(* IEC 61131-3 sources: Caravan/Archiv/12-04-19/Stations/Terminal/HMI/Class/_WeatherForecast (part 2) *)

  for i:=0 to (StrLength - 1) do
    if ((myBuffer[BufferPos - i] >= '0') & (myBuffer[BufferPos - i] <= '9')) then
      case i of
        0: RetValue += TO_DINT((myBuffer[BufferPos - i] - '0') * 1);
        1: RetValue += TO_DINT((myBuffer[BufferPos - i] - '0') * 10);
        2: RetValue += TO_DINT((myBuffer[BufferPos - i] - '0') * 100);
        3: RetValue += TO_DINT((myBuffer[BufferPos - i] - '0') * 1000);
        4: RetValue += TO_DINT((myBuffer[BufferPos - i] - '0') * 10000);
        5: RetValue += TO_DINT((myBuffer[BufferPos - i] - '0') * 100000);
        6: RetValue += TO_DINT((myBuffer[BufferPos - i] - '0') * 1000000);
        7: RetValue += TO_DINT((myBuffer[BufferPos - i] - '0') * 10000000);
        8: RetValue += TO_DINT((myBuffer[BufferPos - i] - '0') * 100000000);
        9: RetValue += TO_DINT((myBuffer[BufferPos - i] - '0') * 1000000000);
      end_case;

    elsif (myBuffer[BufferPos - i] = '-') then    // negate
      RetValue := RetValue * -1;
    elsif ((myBuffer[BufferPos - i] = '.') | (myBuffer[BufferPos - i] = ',')) then    // start again in case of comma
      if ((myBuffer[BufferPos - i+1] - '0') >= 5) then
        RetValue := 1;
      else
        RetValue := 0;
      end_if;
      StrLength -= (i+1);
      i := -1;
      BufferPos := StrLength - 1;
    end_if;

  end_for;

END_FUNCTION

FUNCTION _WeatherForecast::MakeLocalTime
	VAR_INPUT
		pInTime 	: ^CHAR;
		UTC_Offset 	: DINT;
		pRetTime 	: ^CHAR;
	END_VAR

  VAR
  	myTime    : SYSTIME;
  	myDate    : SYSDATE;
    unixtime    : UDINT;
    myTxt : ARRAY [0..20] OF USINT;
  END_VAR

  if ((pInTime <> NIL) & (pRetTime <> NIL)) then

    myTime.wHour   := TO_UINT(CharToDint(pInTime +11, DataLen:=2));
    myTime.wMinute := TO_UINT(CharToDint(pInTime +14, DataLen:=2));
    myTime.wSecond := TO_UINT(CharToDint(pInTime +17, DataLen:=2));
    myTime.wSecond += 1;  // KaiAnd: workaround against UnixTimeStampConvert() bug (2017-10-01 00:00:00 -> 2017-09-31 00:00:00)

    myDate.wYear  := TO_UINT(CharToDint(pInTime +0, DataLen:=4));
    myDate.wMonth := TO_UINT(CharToDint(pInTime +5, DataLen:=2));
    myDate.wDay   := TO_UINT(CharToDint(pInTime +8, DataLen:=2));

    unixtime := SigCLib.UnixTimeStampReconvert(#myDate, #myTime);

    if (UTC_Offset > 0) then
      unixtime += TO_UDINT(UTC_Offset*3600);
    else
      unixtime -= TO_UDINT(UTC_Offset*-1 *3600);
    end_if;

    SigCLib.UnixTimeStampConvert(#myDate, #myTime, unixtime);
    myTime.wSecond -= 1;  // KaiAnd: workaround against UnixTimeStampConvert() bug (2017-10-01 00:00:00 -> 2017-09-31 00:00:00)

    SigCLib.IToA(val:=myDate.wYear, dst:=pRetTime, base:=10);
    SigCLib.StrCat(ps1:=pRetTime, ps2:="-");

    if (myDate.wMonth < 10) then
      SigCLib.StrCat(ps1:=pRetTime, ps2:="0");
    end_if;
    SigCLib.IToA(val:=myDate.wMonth, dst:=#myTxt[0], base:=10);
    SigCLib.StrCat(ps1:=pRetTime, ps2:=#myTxt[0]);
    SigCLib.StrCat(ps1:=pRetTime, ps2:="-");

    if (myDate.wDay < 10) then
      SigCLib.StrCat(ps1:=pRetTime, ps2:="0");
    end_if;
    SigCLib.IToA(val:=myDate.wDay, dst:=#myTxt[0], base:=10);
    SigCLib.StrCat(ps1:=pRetTime, ps2:=#myTxt[0]);
    SigCLib.StrCat(ps1:=pRetTime, ps2:=" ");

    if (myTime.wHour < 10) then
      SigCLib.StrCat(ps1:=pRetTime, ps2:="0");
    end_if;
    SigCLib.IToA(val:=myTime.wHour, dst:=#myTxt[0], base:=10);
    SigCLib.StrCat(ps1:=pRetTime, ps2:=#myTxt[0]);
    SigCLib.StrCat(ps1:=pRetTime, ps2:=":");

    if (myTime.wMinute < 10) then
      SigCLib.StrCat(ps1:=pRetTime, ps2:="0");
    end_if;
    SigCLib.IToA(val:=myTime.wMinute, dst:=#myTxt[0], base:=10);
    SigCLib.StrCat(ps1:=pRetTime, ps2:=#myTxt[0]);
    SigCLib.StrCat(ps1:=pRetTime, ps2:=":");

    if (myTime.wSecond < 10) then
      SigCLib.StrCat(ps1:=pRetTime, ps2:="0");
    end_if;
    SigCLib.IToA(val:=myTime.wSecond, dst:=#myTxt[0], base:=10);
    SigCLib.StrCat(ps1:=pRetTime, ps2:=#myTxt[0]);

  end_if;

END_FUNCTION

FUNCTION _WeatherForecast::MakeSymbolCode
	VAR_INPUT
		pSymbolTxt 	: ^CHAR;
	END_VAR
	VAR_OUTPUT
		SymbolCode 	: INT;
	END_VAR

  if (pSymbolTxt = NIL) then
    SymbolCode := 0;
  else

    // first 2 chars are code, 3rd char is "n" (night) or "d" (day)
    // http://openweathermap.org/weather-conditions
    SymbolCode := TO_INT(CharToDint(pBuffer:=pSymbolTxt, DataLen:=2));
    if ((pSymbolTxt +2)^ = 'n') then
      SymbolCode += 1000;
    elsif ((pSymbolTxt +2)^ = 'd') then
      SymbolCode += 2000;
    end_if;

  end_if;

END_FUNCTION

FUNCTION _WeatherForecast::GetDayMonthWD
	VAR_INPUT
		DayOffset 	: DINT;
		pData 	: ^CHAR;
	END_VAR
  VAR
    DayWork     : DINT;
    DayEntry    : DINT;
    FoundNoDays : DINT;
    i           : DINT;
  END_VAR

  if (pData = NIL) then
    return;
  else
    SigClib.StrCpy(dst0:=pData, src0:=".");
  end_if;

  DayWork := CharToDint(pBuffer:=#WeatherData[0].LocalTime_DateStamp[8], DataLen:=2);
  if (DayWork = 0) then
    return;
  end_if;

  FoundNoDays := 0;
  for i:=0 to (WEATHERFC_XmlEntries-1) do

    DayEntry := CharToDint(pBuffer:=#WeatherData[i].LocalTime_DateStamp[8], DataLen:=2);

    if (DayEntry > 0)then

      if (DayEntry <> DayWork) then
        DayWork := DayEntry;
        FoundNoDays += 1;
      end_if;

      if (FoundNoDays = DayOffset) then
        // timestamp format: "2010-09-31 06:00:00"
        (pData + 0)^ := WeatherData[i].LocalTime_DateStamp[8];
        (pData + 1)^ := WeatherData[i].LocalTime_DateStamp[9];
        (pData + 2)^ := '.';
        (pData + 3)^ := WeatherData[i].LocalTime_DateStamp[5];
        (pData + 4)^ := WeatherData[i].LocalTime_DateStamp[6];
        (pData + 5)^ := 0;
        i := WEATHERFC_XmlEntries;              // escape the loop
      end_if;

    end_if;

  end_for;

END_FUNCTION

FUNCTION _WeatherForecast::GetSymbolCodeWD
	VAR_INPUT
		Hour 	: DINT;
		DayOffset 	: DINT;
	END_VAR
	VAR_OUTPUT
		RetValue 	: DINT;
	END_VAR
  VAR
    DayWork     : DINT;
    DayEntry    : DINT;
    FoundNoDays : DINT;
    i           : DINT;
  END_VAR

  RetValue := 0;
  DayWork := CharToDint(pBuffer:=#WeatherData[0].LocalTime_DateStamp[8], DataLen:=2);
  if (DayWork = 0) then
    return;
  end_if;

  FoundNoDays := 0;
  for i:=0 to (WEATHERFC_XmlEntries-1) do

    DayEntry := CharToDint(pBuffer:=#WeatherData[i].LocalTime_DateStamp[8], DataLen:=2);

    if (DayEntry > 0)then

      if (DayEntry <> DayWork) then
        DayWork := DayEntry;
        FoundNoDays += 1;
      end_if;

      if (FoundNoDays = DayOffset) then
        if (WeatherData[i].LocalTime_fromHH >= Hour) then
          RetValue := WeatherData[i].SymbolCode;  // found the entry!
          i := WEATHERFC_XmlEntries;              // escape the loop
        end_if;
      end_if;

    end_if;

  end_for;

END_FUNCTION

FUNCTION _WeatherForecast::GetWeatherCodeWD
	VAR_INPUT
		Hour 	: DINT;
		DayOffset 	: DINT;
	END_VAR
	VAR_OUTPUT
		RetValue 	: DINT;
	END_VAR
  VAR
    DayWork     : DINT;
    DayEntry    : DINT;
    FoundNoDays : DINT;
    i           : DINT;
  END_VAR

  RetValue := 0;
  DayWork := CharToDint(pBuffer:=#WeatherData[0].LocalTime_DateStamp[8], DataLen:=2);
  if (DayWork = 0) then
    return;
  end_if;

  FoundNoDays := 0;
  for i:=0 to (WEATHERFC_XmlEntries-1) do

    DayEntry := CharToDint(pBuffer:=#WeatherData[i].LocalTime_DateStamp[8], DataLen:=2);

    if (DayEntry > 0)then

      if (DayEntry <> DayWork) then
        DayWork := DayEntry;
        FoundNoDays += 1;
      end_if;

      if (FoundNoDays = DayOffset) then
        if (WeatherData[i].LocalTime_fromHH >= Hour) then
          RetValue := WeatherData[i].SymbolNumber;  // found the entry!
          i := WEATHERFC_XmlEntries;                // escape the loop
        end_if;
      end_if;

    end_if;

  end_for;

END_FUNCTION

FUNCTION _WeatherForecast::GetTempMinWD
	VAR_INPUT
		DayOffset 	: DINT;
	END_VAR
	VAR_OUTPUT
		RetValue 	: DINT;
	END_VAR
  VAR
    DayWork     : DINT;
    DayEntry    : DINT;
    FoundNoDays : DINT;
    myMin       : DINT;
    i           : DINT;
  END_VAR

  RetValue := 0;
  DayWork := CharToDint(pBuffer:=#WeatherData[0].LocalTime_DateStamp[8], DataLen:=2);
  if (DayWork = 0) then
    return;
  end_if;

  FoundNoDays := 0;
  myMin := 9999;
  for i:=0 to (WEATHERFC_XmlEntries-1) do

    DayEntry := CharToDint(pBuffer:=#WeatherData[i].LocalTime_DateStamp[8], DataLen:=2);

    if (DayEntry > 0)then

      if (DayEntry <> DayWork) then
        DayWork := DayEntry;
        FoundNoDays += 1;
      end_if;

      if (FoundNoDays = DayOffset) then
        if (WeatherData[i].TempMin_C < myMin) then
          myMin := WeatherData[i].TempMin_C;
          RetValue := myMin;                // found entry!
        end_if;
      end_if;

    end_if;

  end_for;

END_FUNCTION

FUNCTION _WeatherForecast::GetTempMaxWD
	VAR_INPUT
		DayOffset 	: DINT;
	END_VAR
	VAR_OUTPUT
		RetValue 	: DINT;
	END_VAR
  VAR
    DayWork     : DINT;
    DayEntry    : DINT;
    FoundNoDays : DINT;
    myMax       : DINT;
    i           : DINT;
  END_VAR

  RetValue := 0;
  DayWork := CharToDint(pBuffer:=#WeatherData[0].LocalTime_DateStamp[8], DataLen:=2);
  if (DayWork = 0) then
    return;
  end_if;

  FoundNoDays := 0;
  myMax := -9999;
  for i:=0 to (WEATHERFC_XmlEntries-1) do

    DayEntry := CharToDint(pBuffer:=#WeatherData[i].LocalTime_DateStamp[8], DataLen:=2);

    if (DayEntry > 0)then

      if (DayEntry <> DayWork) then
        DayWork := DayEntry;
        FoundNoDays += 1;
      end_if;

      if (FoundNoDays = DayOffset) then
        if (WeatherData[i].TempMin_C > myMax) then
          myMax := WeatherData[i].TempMax_C;
          RetValue := myMax;                // found entry!
        end_if;
      end_if;

    end_if;

  end_for;

END_FUNCTION

FUNCTION _WeatherForecast::ChkURLchanged
	VAR_OUTPUT
		result 	: DINT;
	END_VAR

	VAR
		newChkSum  : DINT;
    len        : UDINT;
    u 	       : UDINT;
	END_VAR

  result := 0;
  newChkSum := 0;
  len := SigCLib.StrLen(str:=#URL_String[0]);
  for u:=0 to (len -1) do
    newChkSum += URL_String[u];
  end_for;
  if (URL_StringChkSum <> newChkSum) then
    URL_StringChkSum := newChkSum;
    result := 1;
  end_if;

END_FUNCTION

FUNCTION VIRTUAL GLOBAL _WeatherForecast::ProxyAddress::Read
	VAR_OUTPUT
		output (EAX) 	: UDINT;
	END_VAR

	ProxyAddress := Str_ProxyAddress.Data.Read();
	output := ProxyAddress;

END_FUNCTION

FUNCTION VIRTUAL GLOBAL _WeatherForecast::ProxyAddress::Write
	VAR_INPUT
		input (EAX) 	: UDINT;
	END_VAR
	VAR_OUTPUT
		result (EAX) 	: UDINT;
	END_VAR

	ProxyAddress := input;
 	result := (Str_ProxyAddress.Data.Write(ProxyAddress))$UDINT;

END_FUNCTION

FUNCTION VIRTUAL GLOBAL _WeatherForecast::ProxyUser::Read
	VAR_OUTPUT
		output (EAX) 	: UDINT;
	END_VAR

	ProxyUser := Str_ProxyUser.Data.Read();
	output := ProxyUser;

END_FUNCTION

FUNCTION VIRTUAL GLOBAL _WeatherForecast::ProxyUser::Write
	VAR_INPUT
		input (EAX) 	: UDINT;
	END_VAR
	VAR_OUTPUT
		result (EAX) 	: UDINT;
	END_VAR

	ProxyUser := input;
 	result := (Str_ProxyUser.Data.Write(ProxyUser))$UDINT;

END_FUNCTION

FUNCTION VIRTUAL GLOBAL _WeatherForecast::ProxyPassword::Read
	VAR_OUTPUT
		output (EAX) 	: UDINT;
	END_VAR

	ProxyPassword := Str_ProxyPassword.Data.Read();
	output := ProxyPassword;

END_FUNCTION

FUNCTION VIRTUAL GLOBAL _WeatherForecast::ProxyPassword::Write
	VAR_INPUT
		input (EAX) 	: UDINT;
	END_VAR
	VAR_OUTPUT
		result (EAX) 	: UDINT;
	END_VAR

	ProxyPassword := input;
 	result := (Str_ProxyPassword.Data.Write(ProxyPassword))$UDINT;

END_FUNCTION

FUNCTION VIRTUAL GLOBAL _WeatherForecast::ProxyPort::Read
	VAR_OUTPUT
		output (EAX) 	: UDINT;
	END_VAR

	ProxyPort := Str_ProxyPort.Data.Read();
	output := ProxyPort;

END_FUNCTION

FUNCTION VIRTUAL GLOBAL _WeatherForecast::ProxyPort::Write
	VAR_INPUT
		input (EAX) 	: UDINT;
	END_VAR
	VAR_OUTPUT
		result (EAX) 	: UDINT;
	END_VAR

	ProxyPort := input;
 	result := (Str_ProxyPort.Data.Write(ProxyPort))$UDINT;

END_FUNCTION

FUNCTION VIRTUAL GLOBAL _WeatherForecast::WeatherLocName::Read
	VAR_OUTPUT
		output (EAX) 	: UDINT;
	END_VAR

	WeatherLocName := Str_WeatherLocName.Data.Read();
	output := WeatherLocName;

END_FUNCTION

FUNCTION VIRTUAL GLOBAL _WeatherForecast::WeatherLocName::Write
	VAR_INPUT
		input (EAX) 	: UDINT;
	END_VAR
	VAR_OUTPUT
		result (EAX) 	: UDINT;
	END_VAR

	WeatherLocName := input;
 	result := (Str_WeatherLocName.Data.Write(WeatherLocName))$UDINT;

END_FUNCTION

FUNCTION VIRTUAL GLOBAL _WeatherForecast::WeatherLocCountry::Read
	VAR_OUTPUT
		output (EAX) 	: UDINT;
	END_VAR

	WeatherLocCountry := Str_WeatherLocCountry.Data.Read();
	output := WeatherLocCountry;

END_FUNCTION

FUNCTION VIRTUAL GLOBAL _WeatherForecast::WeatherLocCountry::Write
	VAR_INPUT
		input (EAX) 	: UDINT;
	END_VAR
	VAR_OUTPUT
		result (EAX) 	: UDINT;
	END_VAR

	WeatherLocCountry := input;
 	result := (Str_WeatherLocCountry.Data.Write(WeatherLocCountry))$UDINT;

END_FUNCTION

FUNCTION VIRTUAL GLOBAL _WeatherForecast::WeatherUserID::Read
	VAR_OUTPUT
		output (EAX) 	: UDINT;
	END_VAR

	WeatherUserID := Str_WeatherUserID.Data.Read();
	output := WeatherUserID;

END_FUNCTION

FUNCTION VIRTUAL GLOBAL _WeatherForecast::WeatherUserID::Write
	VAR_INPUT
		input (EAX) 	: UDINT;
	END_VAR
	VAR_OUTPUT
		result (EAX) 	: UDINT;
	END_VAR

	WeatherUserID := input;
 	result := (Str_WeatherUserID.Data.Write(WeatherUserID))$UDINT;

END_FUNCTION

FUNCTION VIRTUAL GLOBAL _WeatherForecast::ProxyIsUsed::Write
	VAR_INPUT
		input (EAX) 	: DINT;
	END_VAR
	VAR_OUTPUT
		result (EAX) 	: DINT;
	END_VAR

  if (Status <> -2) then  // if HTTP-client is initialized
    ProxyIsUsed := input;
    result := ProxyIsUsed;
    SetProxy:= TRUE;      // SetOptions(); no method call from a write function v1.01
  end_if;

END_FUNCTION

FUNCTION VIRTUAL GLOBAL _WeatherForecast::Status::Write
	VAR_INPUT
		input (EAX) 	: DINT;
	END_VAR
	VAR_OUTPUT
		result (EAX) 	: DINT;
	END_VAR

  if (Status <> -2) then  // if HTTP-client is initialized
    GetHttpData:= TRUE;
  end_if;

  result := Status;

END_FUNCTION

FUNCTION VIRTUAL GLOBAL _WeatherForecast::WeatherURL::Read
	VAR_OUTPUT
		output (EAX) 	: UDINT;
	END_VAR

	WeatherURL := Str_WeatherURL.Data.Read();
	output := WeatherURL;

END_FUNCTION

FUNCTION VIRTUAL GLOBAL _WeatherForecast::WeatherURL::Write
	VAR_INPUT
		input (EAX) 	: UDINT;
	END_VAR
	VAR_OUTPUT
		result (EAX) 	: UDINT;
	END_VAR

	WeatherURL := input;
 	result := (Str_WeatherURL.Data.Write(WeatherURL))$UDINT;

END_FUNCTION

FUNCTION VIRTUAL GLOBAL _WeatherForecast::Reset_URL::Write
	VAR_INPUT
		input (EAX) 	: DINT;
	END_VAR
	VAR_OUTPUT
		result (EAX) 	: DINT;
	END_VAR

	Reset_URL := input;
 	result := Reset_URL;

  SetWeatherURL();

  Reset_URL := 0;

END_FUNCTION

FUNCTION VIRTUAL GLOBAL _WeatherForecast::WeatherLocID::Read
	VAR_OUTPUT
		output (EAX) 	: UDINT;
	END_VAR

	WeatherLocID := Str_WeatherLocID.Data.Read();
	output := WeatherLocID;

END_FUNCTION

FUNCTION VIRTUAL GLOBAL _WeatherForecast::WeatherLocID::Write
	VAR_INPUT
		input (EAX) 	: UDINT;
	END_VAR
	VAR_OUTPUT
		result (EAX) 	: UDINT;
	END_VAR

	WeatherLocID := input;
	result := (Str_WeatherLocID.Data.Write(WeatherLocID))$UDINT;

END_FUNCTION

FUNCTION VIRTUAL GLOBAL _WeatherForecast::WeatherLocMode::Write
	VAR_INPUT
		input (EAX) 	: DINT;
	END_VAR
	VAR_OUTPUT
		result (EAX) 	: DINT;
	END_VAR

	WeatherLocMode := input;
	result := WeatherLocMode;

END_FUNCTION

FUNCTION VIRTUAL GLOBAL _WeatherForecast::Day1_DD_MM::Read
	VAR_OUTPUT
		output (EAX) 	: UDINT;
	END_VAR

	Day1_DD_MM := Str_Day1_DD_MM.Data.Read();
	output := Day1_DD_MM;

END_FUNCTION

FUNCTION VIRTUAL GLOBAL _WeatherForecast::Day1_DD_MM::Write
	VAR_INPUT
		input (EAX) 	: UDINT;
	END_VAR
	VAR_OUTPUT
		result (EAX) 	: UDINT;
	END_VAR

	Day1_DD_MM := input;
	result := (Str_Day1_DD_MM.Data.Write(Day1_DD_MM))$UDINT;

END_FUNCTION

FUNCTION VIRTUAL GLOBAL _WeatherForecast::Day2_DD_MM::Read
	VAR_OUTPUT
		output (EAX) 	: UDINT;
	END_VAR

	Day2_DD_MM := Str_Day2_DD_MM.Data.Read();
	output := Day2_DD_MM;

END_FUNCTION

FUNCTION VIRTUAL GLOBAL _WeatherForecast::Day2_DD_MM::Write
	VAR_INPUT
		input (EAX) 	: UDINT;
	END_VAR
	VAR_OUTPUT
		result (EAX) 	: UDINT;
	END_VAR

	Day2_DD_MM := input;
	result := (Str_Day2_DD_MM.Data.Write(Day2_DD_MM))$UDINT;

END_FUNCTION

FUNCTION VIRTUAL GLOBAL _WeatherForecast::Day3_DD_MM::Read
	VAR_OUTPUT
		output (EAX) 	: UDINT;
	END_VAR

	Day3_DD_MM := Str_Day3_DD_MM.Data.Read();
	output := Day3_DD_MM;

END_FUNCTION

FUNCTION VIRTUAL GLOBAL _WeatherForecast::Day3_DD_MM::Write
	VAR_INPUT
		input (EAX) 	: UDINT;
	END_VAR
	VAR_OUTPUT
		result (EAX) 	: UDINT;
	END_VAR

	Day3_DD_MM := input;
	result := (Str_Day3_DD_MM.Data.Write(Day3_DD_MM))$UDINT;

END_FUNCTION

FUNCTION VIRTUAL GLOBAL _WeatherForecast::Day4_DD_MM::Read
	VAR_OUTPUT
		output (EAX) 	: UDINT;
	END_VAR

	Day4_DD_MM := Str_Day4_DD_MM.Data.Read();
	output := Day4_DD_MM;

END_FUNCTION

FUNCTION VIRTUAL GLOBAL _WeatherForecast::Day4_DD_MM::Write
	VAR_INPUT
		input (EAX) 	: UDINT;
	END_VAR
	VAR_OUTPUT
		result (EAX) 	: UDINT;
	END_VAR

	Day4_DD_MM := input;
	result := (Str_Day4_DD_MM.Data.Write(Day4_DD_MM))$UDINT;

END_FUNCTION

FUNCTION VIRTUAL GLOBAL _WeatherForecast::Day5_DD_MM::Read
	VAR_OUTPUT
		output (EAX) 	: UDINT;
	END_VAR

	Day5_DD_MM := Str_Day5_DD_MM.Data.Read();
	output := Day5_DD_MM;

END_FUNCTION

FUNCTION VIRTUAL GLOBAL _WeatherForecast::Day5_DD_MM::Write
	VAR_INPUT
		input (EAX) 	: UDINT;
	END_VAR
	VAR_OUTPUT
		result (EAX) 	: UDINT;
	END_VAR

	Day5_DD_MM := input;
	result := (Str_Day5_DD_MM.Data.Write(Day5_DD_MM))$UDINT;

END_FUNCTION

FUNCTION VIRTUAL GLOBAL _WeatherForecast::LastLocationName::Read
	VAR_OUTPUT
		output (EAX) 	: UDINT;
	END_VAR

	LastLocationName := Str_LastLocationName.Data.Read();
	output := LastLocationName;

END_FUNCTION

FUNCTION VIRTUAL GLOBAL _WeatherForecast::LastLocationName::Write
	VAR_INPUT
		input (EAX) 	: UDINT;
	END_VAR
	VAR_OUTPUT
		result (EAX) 	: UDINT;
	END_VAR

	LastLocationName := input;
	result := (Str_LastLocationName.Data.Write(LastLocationName))$UDINT;

END_FUNCTION
